(* IEC 61131-3 sources: Lasal-MCP/examples/SampleSource/LASALScreenAdvancedSolution/LASALScreenAdvancedSolution/LASALScreenAdvacnedSolution/Stations/MachineControl/MachineControl/Class/Tank, 1 file *)

(* ---- Tank.st ---- *)
(*!
<Class
	Name               = "Tank"
	Revision           = "0.0"
	RealtimeTask       = "false"
	CyclicTask         = "false"
	BackgroundTask     = "false"
	Sigmatek           = "false"
	OSInterface        = "false"
	HighPriority       = "false"
	Automatic          = "false"
	UpdateMode         = "Prescan"
	SharedCommandTable = "true"
	Objectsize         = "(484,120)">
	<Channels>
		<Server Name="ActFillLevelVisu" Visualized="true" Initialize="false" WriteProtected="true" Retentive="false"/>
		<Server Name="ClassSvr" Visualized="false" Initialize="false" WriteProtected="true" Retentive="false"/>
		<Server Name="MaxBorder" Visualized="true" Initialize="true" DefValue="45000" WriteProtected="false" Retentive="false"/>
		<Server Name="MinBorder" Visualized="true" Initialize="true" DefValue="10000" WriteProtected="false" Retentive="false"/>
		<Server Name="ShowValue" Visualized="true" Initialize="false" WriteProtected="false" Retentive="false"/>
		<Client Name="ActFillLevel" Required="true" Internal="false"/>
	</Channels>
</Class>
*)
Tank : CLASS
  //Servers:
	ClassSvr 	: SvrChCmd_DINT;
	MinBorder 	: SvrCh_DINT;
	MaxBorder 	: SvrCh_DINT;
	ShowValue 	: SvrCh_DINT;
	ActFillLevelVisu 	: SvrCh_DINT;
  //Clients:
	ActFillLevel 	: CltCh_DINT;
  //Variables:
  //Functions:

	FUNCTION VIRTUAL GLOBAL ActFillLevelVisu::Read
		VAR_OUTPUT
			output (EAX) 	: DINT;
		END_VAR;
  //Tables:
	FUNCTION @STD
		VAR_OUTPUT
			ret_code	: CONFSTATES;
		END_VAR;
	FUNCTION GLOBAL TAB @CT_;
END_CLASS;

FUNCTION VIRTUAL GLOBAL Tank::ActFillLevelVisu::Read
	VAR_OUTPUT
		output (EAX) 	: DINT;
	END_VAR

  ActFillLevel := ActFillLevel.Read();

	ActFillLevelVisu := ActFillLevel;

	output := ActFillLevelVisu;

END_FUNCTION
